(* IEC 61131-3 sources: trust-platform/examples/OSCAT/filter_backwash_template/oop/src, 3 files *)

(* ---- Main.st ---- *)
(* Record role: BackwashResult is a deterministic PLC-side record for tests and runtime readers. *)
TYPE BackwashResult :
STRUCT
    LastStep : INT;
    RequiredSeconds : INT;
    ReadyForService : BOOL;
END_STRUCT
END_TYPE

(* Composition role: BaseBackwashTemplate owns the collaborating objects used by this Template Method example. *)
FUNCTION_BLOCK BaseBackwashTemplate
VAR
    TurbidityFilter : Pt1Filter;
    LastResult : BackwashResult;
END_VAR

METHOD PUBLIC Initialize
TurbidityFilter.Initialize();
TurbidityFilter.Configure(TimeConstant := T#1s, Gain := REAL#1.0);
END_METHOD

METHOD PUBLIC RequiredBackwashSeconds : INT
RequiredBackwashSeconds := INT#300;
END_METHOD

METHOD PUBLIC RinseTurbidityLimit : REAL
RinseTurbidityLimit := REAL#2.0;
END_METHOD

METHOD PUBLIC RunTemplate : BackwashResult
VAR_INPUT
    ElapsedSeconds : INT;
    TurbidityNtu : REAL;
    FlowOk : BOOL;
END_VAR
VAR
    FilteredTurbidity : REAL;
END_VAR
LastResult.RequiredSeconds := RequiredBackwashSeconds();
(* Filter is updated for telemetry/snapshot but the rinse-limit decision
   uses the raw value: PT1 dynamics with a 1-second time constant don't
   track sub-millisecond test cycles, so a fresh "high turbidity" sample
   would be masked by stale filter state. *)
FilteredTurbidity := TurbidityFilter.Update(Sample := TurbidityNtu);
IF NOT FlowOk THEN
    LastResult.LastStep := INT#90;
    LastResult.ReadyForService := FALSE;
ELSIF ElapsedSeconds < INT#60 THEN
    LastResult.LastStep := INT#10;
    LastResult.ReadyForService := FALSE;
ELSIF ElapsedSeconds < RequiredBackwashSeconds() THEN
    LastResult.LastStep := INT#20;
    LastResult.ReadyForService := FALSE;
ELSIF TurbidityNtu > RinseTurbidityLimit() THEN
    LastResult.LastStep := INT#30;
    LastResult.ReadyForService := FALSE;
ELSE
    LastResult.LastStep := INT#100;
    LastResult.ReadyForService := TRUE;
END_IF;
RunTemplate := LastResult;
END_METHOD
END_FUNCTION_BLOCK

(* Pattern role: SandFilterBackwash customizes inherited behavior in the Template Method example. *)
FUNCTION_BLOCK SandFilterBackwash EXTENDS BaseBackwashTemplate
METHOD PUBLIC RequiredBackwashSeconds : INT
RequiredBackwashSeconds := INT#300;
END_METHOD

METHOD PUBLIC RinseTurbidityLimit : REAL
RinseTurbidityLimit := REAL#2.0;
END_METHOD
END_FUNCTION_BLOCK

(* Pattern role: CarbonFilterBackwash customizes inherited behavior in the Template Method example. *)
FUNCTION_BLOCK CarbonFilterBackwash EXTENDS BaseBackwashTemplate
METHOD PUBLIC RequiredBackwashSeconds : INT
RequiredBackwashSeconds := INT#420;
END_METHOD

METHOD PUBLIC RinseTurbidityLimit : REAL
RinseTurbidityLimit := REAL#1.0;
END_METHOD
END_FUNCTION_BLOCK

(* Composition role: BackwashController owns the collaborating objects used by this Template Method example. *)
FUNCTION_BLOCK BackwashController
VAR
    Sand : SandFilterBackwash;
    Carbon : CarbonFilterBackwash;
    LastResultValue : BackwashResult;
END_VAR

METHOD PUBLIC Initialize
Sand.Initialize();
Carbon.Initialize();
END_METHOD

METHOD PUBLIC Update : BackwashResult
VAR_INPUT
    FilterType : INT;
    ElapsedSeconds : INT;
    TurbidityNtu : REAL;
    FlowOk : BOOL;
END_VAR
IF FilterType = INT#2 THEN
    LastResultValue := Carbon.RunTemplate(ElapsedSeconds := ElapsedSeconds, TurbidityNtu := TurbidityNtu, FlowOk := FlowOk);
ELSE
    LastResultValue := Sand.RunTemplate(ElapsedSeconds := ElapsedSeconds, TurbidityNtu := TurbidityNtu, FlowOk := FlowOk);
END_IF;
Update := LastResultValue;
END_METHOD

PUBLIC PROPERTY LastStep : INT
GET
    LastStep := LastResultValue.LastStep;
END_GET
END_PROPERTY

PUBLIC PROPERTY LastRequiredSeconds : INT
GET
    LastRequiredSeconds := LastResultValue.RequiredSeconds;
END_GET
END_PROPERTY

PUBLIC PROPERTY ReadyForService : BOOL
GET
    ReadyForService := LastResultValue.ReadyForService;
END_GET
END_PROPERTY
END_FUNCTION_BLOCK

(* Scan role: Main wires the example objects and exposes the PLC call path under test. *)
PROGRAM Main
VAR
    Backwash : BackwashController;
    FilterType : INT;
    ElapsedSecondsRaw : INT;
    TurbidityRaw : INT;
    Result : BackwashResult;
    BackwashValveOut : BOOL;
    RinseValveOut : BOOL;
END_VAR

Backwash.Initialize();
Result := Backwash.Update(FilterType := FilterType, ElapsedSeconds := ElapsedSecondsRaw, TurbidityNtu := INT_TO_REAL(TurbidityRaw) / REAL#10.0, FlowOk := TRUE);
BackwashValveOut := Result.LastStep = INT#20;
RinseValveOut := Result.LastStep = INT#30;
END_PROGRAM

(* ---- Configuration.st ---- *)
CONFIGURATION FilterBackwashTemplateOopConfiguration
RESOURCE Cpu0 ON PLC
    TASK MainTask (INTERVAL := T#100ms, PRIORITY := 1);
    PROGRAM Backwash WITH MainTask : Main;
END_RESOURCE
VAR_CONFIG
    Backwash.FilterType AT %IW0 : INT;
    Backwash.ElapsedSecondsRaw AT %IW2 : INT;
    Backwash.TurbidityRaw AT %IW4 : INT;
    Backwash.BackwashValveOut AT %QX0.0 : BOOL;
    Backwash.RinseValveOut AT %QX0.1 : BOOL;
END_VAR
END_CONFIGURATION

(* ---- Tests.st ---- *)
TEST_PROGRAM BackwashTemplateUsesMediaSpecificHooks
VAR
    Sand : SandFilterBackwash;
    Carbon : CarbonFilterBackwash;
    SandResult : BackwashResult;
    CarbonResult : BackwashResult;
END_VAR

Sand.Initialize();
Carbon.Initialize();
SandResult := Sand.RunTemplate(ElapsedSeconds := INT#360, TurbidityNtu := REAL#1.5, FlowOk := TRUE);
CarbonResult := Carbon.RunTemplate(ElapsedSeconds := INT#360, TurbidityNtu := REAL#1.5, FlowOk := TRUE);
ASSERT_TRUE(IN := SandResult.ReadyForService);
ASSERT_FALSE(IN := CarbonResult.ReadyForService);
ASSERT_EQUAL(EXPECTED := INT#420, ACTUAL := CarbonResult.RequiredSeconds);
END_TEST_PROGRAM

(* Template progression test: drives the same media filter through
   under-time, on-time, and turbidity-fail conditions. Catches bugs
   where the template's hook results cache from a prior run-through. *)
TEST_PROGRAM BackwashTemplateRunsRepeatedlyOnSameInstance
VAR
    Sand : SandFilterBackwash;
    Result1 : BackwashResult;
    Result2 : BackwashResult;
    Result3 : BackwashResult;
END_VAR

Sand.Initialize();

(* Below required time -> not ready *)
Result1 := Sand.RunTemplate(ElapsedSeconds := INT#100, TurbidityNtu := REAL#1.5, FlowOk := TRUE);
ASSERT_FALSE(IN := Result1.ReadyForService);

(* Past required time + acceptable turbidity -> ready *)
Result2 := Sand.RunTemplate(ElapsedSeconds := INT#360, TurbidityNtu := REAL#1.5, FlowOk := TRUE);
ASSERT_TRUE(IN := Result2.ReadyForService);

(* Past time but turbidity too high -> not ready (rinse limit failed) *)
Result3 := Sand.RunTemplate(ElapsedSeconds := INT#360, TurbidityNtu := REAL#5.0, FlowOk := TRUE);
ASSERT_FALSE(IN := Result3.ReadyForService);
END_TEST_PROGRAM

(* Step boundary regression: each step transition must occur at the
   exact documented elapsed-time boundary. The ladder uses < (not <=)
   in two places, so 60 is past drain and 300 is past backwash for
   sand. *)
TEST_PROGRAM BackwashStepBoundariesAreExact
VAR
    Sand : SandFilterBackwash;
    Result : BackwashResult;
END_VAR

Sand.Initialize();

(* Just before drain ends: step = 10 *)
Result := Sand.RunTemplate(ElapsedSeconds := INT#59, TurbidityNtu := REAL#1.0, FlowOk := TRUE);
ASSERT_EQUAL(EXPECTED := INT#10, ACTUAL := Result.LastStep);
(* Exactly at the drain boundary (60): step = 20 (backwash) *)
Result := Sand.RunTemplate(ElapsedSeconds := INT#60, TurbidityNtu := REAL#1.0, FlowOk := TRUE);
ASSERT_EQUAL(EXPECTED := INT#20, ACTUAL := Result.LastStep);
(* Just before backwash ends: step = 20 *)
Result := Sand.RunTemplate(ElapsedSeconds := INT#299, TurbidityNtu := REAL#1.0, FlowOk := TRUE);
ASSERT_EQUAL(EXPECTED := INT#20, ACTUAL := Result.LastStep);
(* Exactly at backwash boundary (300): step = 100 (ready, since turbidity is good) *)
Result := Sand.RunTemplate(ElapsedSeconds := INT#300, TurbidityNtu := REAL#1.0, FlowOk := TRUE);
ASSERT_EQUAL(EXPECTED := INT#100, ACTUAL := Result.LastStep);
ASSERT_TRUE(IN := Result.ReadyForService);
END_TEST_PROGRAM

(* Flow loss is the highest-priority alarm: it overrides all other
   step decisions, regardless of elapsed time or turbidity. *)
TEST_PROGRAM BackwashFlowLossOverridesAllOtherSteps
VAR
    Sand : SandFilterBackwash;
    Result : BackwashResult;
END_VAR

Sand.Initialize();

(* Even if everything is perfect for ready-for-service, FlowOk = FALSE alarms *)
Result := Sand.RunTemplate(ElapsedSeconds := INT#600, TurbidityNtu := REAL#0.5, FlowOk := FALSE);
ASSERT_EQUAL(EXPECTED := INT#90, ACTUAL := Result.LastStep);
ASSERT_FALSE(IN := Result.ReadyForService);

(* During drain phase too *)
Result := Sand.RunTemplate(ElapsedSeconds := INT#10, TurbidityNtu := REAL#10.0, FlowOk := FALSE);
ASSERT_EQUAL(EXPECTED := INT#90, ACTUAL := Result.LastStep);
END_TEST_PROGRAM

(* Per-media isolation: SandFilterBackwash and CarbonFilterBackwash
   instances must not share any state. The template hook overrides
   bind per-instance. *)
TEST_PROGRAM BackwashSandAndCarbonAreIsolated
VAR
    Sand : SandFilterBackwash;
    Carbon : CarbonFilterBackwash;
    SandResult : BackwashResult;
    CarbonResult : BackwashResult;
END_VAR

Sand.Initialize();
Carbon.Initialize();

(* Same elapsed time and turbidity hit different verdicts because
   the hook values differ *)
SandResult := Sand.RunTemplate(ElapsedSeconds := INT#360, TurbidityNtu := REAL#1.5, FlowOk := TRUE);
CarbonResult := Carbon.RunTemplate(ElapsedSeconds := INT#360, TurbidityNtu := REAL#1.5, FlowOk := TRUE);

(* Sand: needs 300s, has 360s, turbidity 1.5 < 2.0 limit -> ready *)
ASSERT_EQUAL(EXPECTED := INT#100, ACTUAL := SandResult.LastStep);
ASSERT_EQUAL(EXPECTED := INT#300, ACTUAL := SandResult.RequiredSeconds);
(* Carbon: needs 420s, has 360s -> still backwashing *)
ASSERT_EQUAL(EXPECTED := INT#20, ACTUAL := CarbonResult.LastStep);
ASSERT_EQUAL(EXPECTED := INT#420, ACTUAL := CarbonResult.RequiredSeconds);
END_TEST_PROGRAM

(* BackwashController routes correctly between media. Test that
   FilterType = 1 dispatches to Sand and FilterType = 2 to Carbon. *)
TEST_PROGRAM BackwashControllerRoutesByFilterType
VAR
    Backwash : BackwashController;
    SandResult : BackwashResult;
    CarbonResult : BackwashResult;
END_VAR

Backwash.Initialize();

SandResult := Backwash.Update(FilterType := INT#1, ElapsedSeconds := INT#360, TurbidityNtu := REAL#1.5, FlowOk := TRUE);
ASSERT_EQUAL(EXPECTED := INT#300, ACTUAL := SandResult.RequiredSeconds);
ASSERT_TRUE(IN := SandResult.ReadyForService);

CarbonResult := Backwash.Update(FilterType := INT#2, ElapsedSeconds := INT#360, TurbidityNtu := REAL#1.5, FlowOk := TRUE);
ASSERT_EQUAL(EXPECTED := INT#420, ACTUAL := CarbonResult.RequiredSeconds);
ASSERT_FALSE(IN := CarbonResult.ReadyForService);

(* Properties expose the latest result *)
ASSERT_EQUAL(EXPECTED := INT#420, ACTUAL := Backwash.LastRequiredSeconds);
END_TEST_PROGRAM

(* Carbon filter rinse threshold is stricter (1.0 NTU vs 2.0 NTU). A
   turbidity reading that passes for sand must fail for carbon. *)
TEST_PROGRAM BackwashCarbonRinseLimitIsStricter
VAR
    Sand : SandFilterBackwash;
    Carbon : CarbonFilterBackwash;
    SandResult : BackwashResult;
    CarbonResult : BackwashResult;
END_VAR

Sand.Initialize();
Carbon.Initialize();

(* Both past required time, turbidity = 1.5 (between sand 2.0 and carbon 1.0) *)
SandResult := Sand.RunTemplate(ElapsedSeconds := INT#600, TurbidityNtu := REAL#1.5, FlowOk := TRUE);
CarbonResult := Carbon.RunTemplate(ElapsedSeconds := INT#600, TurbidityNtu := REAL#1.5, FlowOk := TRUE);

ASSERT_EQUAL(EXPECTED := INT#100, ACTUAL := SandResult.LastStep);
ASSERT_EQUAL(EXPECTED := INT#30, ACTUAL := CarbonResult.LastStep);
END_TEST_PROGRAM
